PROGRAM motor_ladder
VAR
END_VAR

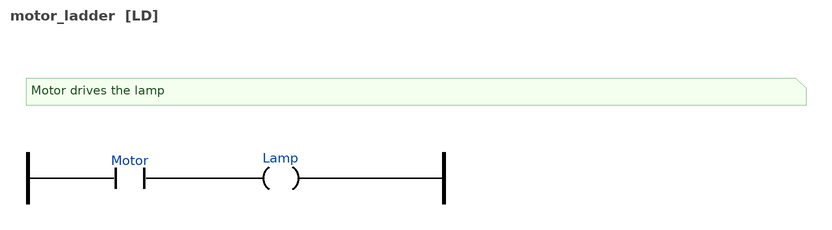
(* LD diagram, written out as Structured Text *)
(* Motor drives the lamp *)
Lamp := Motor;
END_PROGRAM
